(* PLC project RobotLibrarySysDep, Rexroth ctrlX PLC Engineering ctrlX PLC 3.6.3, author Thorsten Brach *)
(* stored: creationDateTime 2026-09-19T14:40:47.4551079, version 0.0.0.2, modificationDateTime 2026-09-19T14:40:11.6627075, organization Thorsten Brach *)
(* SRCI Robot Library System Dependencies *)

FUNCTION SysDepMemCmp : DINT
// ------------------------------------------------------------------------- 
//  SRCI Robot Library System Dependencies                                               
// ------------------------------------------------------------------------- 
//                                                                           
//  Object:      SysDepMemCmp                                       
//  Author:      Thorsten Brach                                                
//  Date:        2024-12-21
//
//  Description:                                              
//    System specific implementation of the memory compare function 
//                                                                           
//  Copyright: 
//    (C) 2024 Thorsten Brach. All rights reserved                                                                                                                                            
//             Licensed under the MIT License.
//                                                                           
//  Disclaimer:                                                                           
//    This project is provided without any guarantee and can be used for   
//    private and commercial purposes. Any use is at the user’s 
//    own risk and responsibility.
//
// -------------------------------------------------------------------------
VAR_INPUT
  /// Pointer to 1st memory area to be compared with the 2nd memory area
  pData1 : POINTER TO BYTE;
  /// Pointer to 2nd memory area to be compared with the 1st memory area
  pData2 : POINTER TO BYTE;
  /// Amount of bytes to be compared
  DataLen : UDINT;
END_VAR

            SysDepMemCmp := SysMemCmp( pBuffer1 := pData1, pBuffer2 := pData2, udiCount := DataLen );

          
END_FUNCTION

FUNCTION SysDepMemCpy : UDINT
// ------------------------------------------------------------------------- 
//  SRCI Robot Library System Dependencies                                               
// ------------------------------------------------------------------------- 
//                                                                           
//  Object:      SysDepMemCpy                                       
//  Author:      Thorsten Brach                                                
//  Date:        2024-12-21
//
//  Description:                                              
//    System specific implementation of the memory copy function 
//                                                                           
//  Copyright: 
//    (C) 2024 Thorsten Brach. All rights reserved                                                                                                                                            
//             Licensed under the MIT License.
//                                                                           
//  Disclaimer:                                                                           
//    This project is provided without any guarantee and can be used for   
//    private and commercial purposes. Any use is at the user’s 
//    own risk and responsibility.
//
// -------------------------------------------------------------------------
VAR_INPUT
  /// Pointer to memory address to be copied to (target)
  pDest : POINTER TO BYTE;
  /// Pointer to memory address to be copied from (source)
  pSrc : POINTER TO BYTE;
  /// Amount of bytes to be copied
  DataLen : UDINT;
END_VAR

            SysMemCpy( pDest := pDest, pSrc := pSrc, udiCount := DataLen );


          
END_FUNCTION

FUNCTION SysDepMemSet : UDINT
// ------------------------------------------------------------------------- 
//  SRCI Robot Library System Dependencies                                               
// ------------------------------------------------------------------------- 
//                                                                           
//  Object:      SysDepMemSet                                       
//  Author:      Thorsten Brach                                                
//  Date:        2024-12-21
//
//  Description:                                              
//    System specific implementation of the memory set function 
//                                                                           
//  Copyright: 
//    (C) 2024 Thorsten Brach. All rights reserved                                                                                                                                            
//             Licensed under the MIT License.
//                                                                           
//  Disclaimer:                                                                           
//    This project is provided without any guarantee and can be used for   
//    private and commercial purposes. Any use is at the user’s 
//    own risk and responsibility.
//
// -------------------------------------------------------------------------
VAR_INPUT
  /// Pointer to memory address to be filled (target)
  pDest : POINTER TO BYTE;
  /// Value with which the memory is to be initialized
  Value : BYTE;
  /// Amount of bytes to be initialized in the memory block
  DataLen : UDINT;
END_VAR

            SysMemSet( pDest := pDest, udiValue := Value, udiCount := DataLen );
          
END_FUNCTION

FUNCTION SysDepIsValidLReal : BOOL
// ------------------------------------------------------------------------- 
//  SRCI Robot Library System Dependencies                                               
// ------------------------------------------------------------------------- 
//                                                                           
//  Object:      SysDepIsValidLReal                                       
//  Author:      Thorsten Brach                                                
//  Date:        2025-03-04
//
//  Description:                                              
//    System specific implementation of the memory compare function 
//                                                                           
//  Copyright: 
//    (C) 2025 Thorsten Brach. All rights reserved                                                                                                                                            
//             Licensed under the MIT License.
//                                                                           
//  Disclaimer:                                                                           
//    This project is provided without any guarantee and can be used for   
//    private and commercial purposes. Any use is at the user’s 
//    own risk and responsibility.
//
// -------------------------------------------------------------------------
VAR_INPUT
  /// Real value to validate
  Value : LREAL;
END_VAR

            SysDepIsValidLReal := FPU.IsLRealNumber(Value);
          
END_FUNCTION

FUNCTION SysDepIsValidReal : BOOL
// ------------------------------------------------------------------------- 
//  SRCI Robot Library System Dependencies                                               
// ------------------------------------------------------------------------- 
//                                                                           
//  Object:      SysDepIsValidReal                                       
//  Author:      Thorsten Brach                                                
//  Date:        2025-03-04
//
//  Description:                                              
//    System specific implementation of the memory compare function 
//                                                                           
//  Copyright: 
//    (C) 2025 Thorsten Brach. All rights reserved                                                                                                                                            
//             Licensed under the MIT License.
//                                                                           
//  Disclaimer:                                                                           
//    This project is provided without any guarantee and can be used for   
//    private and commercial purposes. Any use is at the user’s 
//    own risk and responsibility.
//
// -------------------------------------------------------------------------
VAR_INPUT
  /// Real value to validate
  Value : REAL;
END_VAR

            SysDepIsValidReal := FPU.IsRealNumber(Value);
          
END_FUNCTION
